(* IEC 61131-3 sources: KinematicsSimulation/crates/sim-opcua/examples/plc/twincat, 3 files *)

(* ---- sim_cycle.st ---- *)
(*
    A PLC cycle against the KinematicsSimulation link (sim-opcua), for TwinCAT 3 with TF6100 (library
    Tc3_PLCopen_OpcUa). Uses SIM_Access, SIM_MC_Power and SIM_MC_MoveAbsolute from sim_plcopen.st in this folder.

    NOT COMPILED: TwinCAT needs a Beckhoff account to download, so it was not built. The names were checked on
    14 November 2026 against Beckhoff Infosys (TF6100 TwinCAT 3 OPC UA Client, documentation 1.3.0 of 8 April 2026)
    and Beckhoff's TF6100_Samples on GitHub; what those do not settle is marked "CHECK".

    PRG_SimCycle:
      - connects with Basic256Sha256 SignAndEncrypt (or None, see bSecure), optionally with user name and password;
      - finds the namespace index from the URI 'urn:kinematics-simulation';
      - gets the node handles of the position and following error of one axis once and reads both every cycle,
        with the handles kept (one round trip per read; a read is started again as soon as the last one is done);
      - powers the axis (MC_Power), moves it with MC_MoveAbsolute, then writes a path and runs it
        (command.path, command.run_path) and waits until status.busy falls;
      - keeps the largest following error seen, switches off and disconnects.
    Run it in a task of 10 ms; sim-opcua then reports the task's write and read intervals (status.client_*).

    Data types as sim-opcua serves them (docs/plc.md, "Node ids and data types"): Double -> LREAL, Boolean -> BOOL,
    UInt16 -> UINT, Int32 -> DINT, UInt64 -> ULINT, String -> STRING. A PLC variable of another type (REAL for a
    Double) makes UA_Read fail with a type mismatch.
*)

FUNCTION_BLOCK SIM_CyclicRead
(* Reads one LREAL variable over and over through a node handle that is got once. *)
VAR_INPUT
    bEnable     : BOOL;
    hConnection : DWORD;
    nNamespace  : UINT;
    sNode       : STRING(255);
END_VAR
VAR_OUTPUT
    fValue  : LREAL;
    nReads  : UDINT;     (* reads done *)
    bError  : BOOL;
    nErrorID : DWORD;
END_VAR
VAR
    fbGetHandle : UA_NodeGetHandle;
    fbRead      : UA_Read;
    fbRelease   : UA_NodeReleaseHandle;
    stNodeID    : ST_UANodeID;
    stInfo      : ST_UANodeAdditionalInfo;
    hNode       : DWORD;
    nStep       : INT;
END_VAR

CASE nStep OF
0:  IF bEnable THEN
        stNodeID.nNamespaceIndex := nNamespace;
        stNodeID.sIdentifier := sNode;
        stNodeID.eIdentifierType := eUAIdentifierType_String;
        stInfo.eAttributeID := eUAAI_Value;   (* the Value attribute, 13 *)
        bError := FALSE; nErrorID := 0;
        nStep := 1;
    END_IF
1:  fbGetHandle(Execute := TRUE, ConnectionHdl := hConnection, NodeID := stNodeID);
    IF fbGetHandle.Done THEN
        hNode := fbGetHandle.NodeHdl; fbGetHandle(Execute := FALSE); nStep := 2;
    ELSIF fbGetHandle.Error THEN
        nErrorID := fbGetHandle.ErrorID; fbGetHandle(Execute := FALSE); bError := TRUE; nStep := 9;
    END_IF
2:  (* one read; once it is done the next starts in the same cycle, so a read that returns within a cycle runs
       every cycle *)
    fbRead(Execute := TRUE, ConnectionHdl := hConnection, NodeHdl := hNode, stNodeAddInfo := stInfo,
           cbData := SIZEOF(fValue), pVariable := ADR(fValue));
    IF fbRead.Done OR fbRead.Error THEN
        IF fbRead.Error THEN bError := TRUE; nErrorID := fbRead.ErrorID; ELSE nReads := nReads + 1; END_IF
        fbRead(Execute := FALSE);
        IF bEnable THEN
            fbRead(Execute := TRUE, ConnectionHdl := hConnection, NodeHdl := hNode, stNodeAddInfo := stInfo,
                   cbData := SIZEOF(fValue), pVariable := ADR(fValue));
        ELSE
            nStep := 3;
        END_IF
    END_IF
3:  fbRelease(Execute := TRUE, ConnectionHdl := hConnection, NodeHdl := hNode);
    IF fbRelease.Done OR fbRelease.Error THEN fbRelease(Execute := FALSE); nStep := 0; END_IF
9:  IF NOT bEnable THEN nStep := 0; END_IF
END_CASE
END_FUNCTION_BLOCK

PROGRAM PRG_SimCycle
VAR
    sServerUrl   : STRING(255) := 'opc.tcp://127.0.0.1:4840';   (* sim-opcua on the same PC *)
    bSecure      : BOOL := TRUE;                                 (* FALSE: SecurityPolicy None *)
    sUser        : STRING(63) := '';                             (* empty: anonymous; else as sim-opcua --user *)
    sPassword    : STRING(63) := '';
    sAxis        : STRING(31) := 'x';                            (* an axis id of the simulated machine *)
    fTarget      : LREAL := 0.4;                                 (* m, inside the axis range *)
    (* The path in the text of a path file, one piece per line ($N), one position per axis (here x and z of the
       T-gantry, which starts at x 0.1, z 0.35). *)
    sPath        : STRING(255) := 'line,0.4,0.25$Nline,0.1,0.25$Nline,0.1,0.35';
    (* sim-opcua counts every Read request: two reads a cycle show as intervals of half a cycle. FALSE reads the
       position alone, one request a cycle, so status.client_read_* give the task's cycle and jitter. *)
    bReadFollowingError : BOOL := TRUE;

    fbConnect    : UA_Connect;
    fbNamespace  : UA_GetNamespaceIndex;
    fbDisconnect : UA_Disconnect;
    stSession    : ST_UASessionConnectInfo;
    hConnection  : DWORD;
    nNamespace   : UINT;
    fbPower      : SIM_MC_Power;
    fbMove       : SIM_MC_MoveAbsolute;
    fbWrite      : SIM_Access;
    fbBusy       : SIM_Access;
    fbPosition   : SIM_CyclicRead;
    fbError      : SIM_CyclicRead;
    bTrue        : BOOL := TRUE;
    bBusy        : BOOL;
    bBusySeen    : BOOL;
    fLargestError : LREAL;   (* m, the largest following error read *)
    nStep        : INT;
END_VAR

CASE nStep OF
0:  stSession.sApplicationName := 'TwinCAT sim client';
    stSession.eTransportProfileUri := eUATransportProfileUri_UATcp;
    stSession.tSessionTimeout := T#60S;
    IF bSecure THEN
        (* TF6100 creates its own self-signed client certificate on its first start, in its PKI folder
           (%TcInstallDir%\3.1\Target\OpcUa\Client\PKI for client 2.x, %ProgramData%\Beckhoff\TF6100-OPC-UA\
           TcOpcUaClient\PKI for 1.x; Infosys "Application directories"). sim-opcua refuses it once and stores it in
           pki/rejected; move it to pki/trusted, or start sim-opcua with --trust-all while commissioning. TF6100
           likewise puts the server's certificate into its own rejected folder on the first attempt: move it to
           trusted there. *)
        stSession.eSecurityMode := eUASecurityMsgMode_Sign_Encrypt;
        stSession.eSecurityPolicyUri := eUASecurityPolicy_Basic256Sha256;
    ELSE
        stSession.eSecurityMode := eUASecurityMsgMode_None;
        stSession.eSecurityPolicyUri := eUASecurityPolicy_None;
    END_IF
    IF LEN(sUser) > 0 THEN
        stSession.stUserIdentTokenType.eUserIdentTokenType := eUAUITT_Username;
        stSession.stUserIdentTokenType.sTokenParam1 := sUser;
        stSession.stUserIdentTokenType.sTokenParam2 := sPassword;
    END_IF
    fbConnect(Execute := TRUE, ServerURL := sServerUrl, SessionConnectInfo := stSession, Timeout := T#5S);
    IF fbConnect.Done THEN hConnection := fbConnect.ConnectionHdl; fbConnect(Execute := FALSE); nStep := 10;
    ELSIF fbConnect.Error THEN fbConnect(Execute := FALSE); nStep := 900; END_IF
10: fbNamespace(Execute := TRUE, ConnectionHdl := hConnection, NamespaceUri := 'urn:kinematics-simulation', Timeout := T#5S);
    IF fbNamespace.Done THEN nNamespace := fbNamespace.NamespaceIndex; fbNamespace(Execute := FALSE); nStep := 20;
    ELSIF fbNamespace.Error THEN fbNamespace(Execute := FALSE); nStep := 900; END_IF
20: (* enable the drives *)
    fbPower.Enable := TRUE;
    IF fbPower.Status THEN nStep := 30; END_IF
30: (* MC_MoveAbsolute *)
    fbMove.Position := fTarget; fbMove.Velocity := 0.5; fbMove.Acceleration := 5.0; fbMove.Deceleration := 5.0;
    fbMove.Jerk := 100.0;
    fbMove.Execute := TRUE;
    IF fbMove.Done THEN fbMove.Execute := FALSE; nStep := 40;
    ELSIF fbMove.Error OR fbMove.CommandAborted THEN nStep := 900; END_IF
40: (* the path: its text, then command.run_path *)
    fbWrite(bExecute := FALSE);
    fbWrite(bExecute := TRUE, hConnection := hConnection, nNamespace := nNamespace, sNode := 'command.path',
            bWrite := TRUE, pData := ADR(sPath), cbData := LEN(sPath));
            (* CHECK: UA_Write documents cbData only as the size of the values to write; whether a STRING takes
               LEN (without the terminating null) or SIZEOF (the whole declared buffer) it does not say. *)
    nStep := 41;
41: fbWrite(bExecute := TRUE);
    IF fbWrite.bDone THEN nStep := 42; ELSIF fbWrite.bError THEN nStep := 900; END_IF
42: fbWrite(bExecute := FALSE);
    fbWrite(bExecute := TRUE, hConnection := hConnection, nNamespace := nNamespace, sNode := 'command.run_path',
            bWrite := TRUE, pData := ADR(bTrue), cbData := SIZEOF(bTrue));
    nStep := 43;
43: fbWrite(bExecute := TRUE);
    IF fbWrite.bDone THEN bBusySeen := FALSE; nStep := 50; ELSIF fbWrite.bError THEN nStep := 900; END_IF
50: (* poll status.busy until the path is over: it rises within a loop cycle or two and falls at the end *)
    fbBusy(bExecute := FALSE);
    fbBusy(bExecute := TRUE, hConnection := hConnection, nNamespace := nNamespace, sNode := 'status.busy',
           bWrite := FALSE, pData := ADR(bBusy), cbData := SIZEOF(bBusy));
    nStep := 51;
51: fbBusy(bExecute := TRUE);
    IF fbBusy.bDone THEN
        IF bBusy THEN bBusySeen := TRUE; nStep := 50;
        ELSIF bBusySeen THEN nStep := 60;
        ELSE nStep := 50; END_IF
    ELSIF fbBusy.bError THEN nStep := 900; END_IF
60: (* switch off and disconnect *)
    fbPower.Enable := FALSE;
    IF NOT fbPower.Status THEN nStep := 70; END_IF
70: fbDisconnect(Execute := TRUE, ConnectionHdl := hConnection, Timeout := T#5S);
    IF fbDisconnect.Done OR fbDisconnect.Error THEN fbDisconnect(Execute := FALSE); nStep := 100; END_IF
100: ; (* finished: fLargestError holds the largest following error *)
900: ; (* error: look at the blocks' ErrorID and at status.refused on the server *)
END_CASE

(* every cycle from the namespace on: position and following error of the axis *)
fbPosition(bEnable := nStep >= 20 AND nStep < 70, hConnection := hConnection, nNamespace := nNamespace,
           sNode := CONCAT(CONCAT('signal.axis.', sAxis), '.position'));
fbError(bEnable := bReadFollowingError AND nStep >= 20 AND nStep < 70, hConnection := hConnection, nNamespace := nNamespace,
        sNode := CONCAT(CONCAT('signal.axis.', sAxis), '.following_error'));
IF ABS(fbError.fValue) > fLargestError THEN fLargestError := ABS(fbError.fValue); END_IF

IF nStep >= 20 AND nStep < 70 THEN
    fbPower(hConnection := hConnection, nNamespace := nNamespace, sAxis := sAxis);
    fbMove(hConnection := hConnection, nNamespace := nNamespace, sAxis := sAxis);
END_IF
END_PROGRAM

(* ---- sim_plcopen.st ---- *)
(*
    PLCopen motion over OPC UA to the KinematicsSimulation link (sim-opcua), for TwinCAT 3.
    Library: Tc3_PLCopen_OpcUa (add it in the PLC project's References).

    NOT COMPILED: TwinCAT needs a Beckhoff account to download, so this file was not built. The names were checked
    on 14 November 2026 against Beckhoff Infosys (TF6100 TwinCAT 3 OPC UA Client, documentation 1.3.0 of
    8 April 2026) and Beckhoff's TF6100_Samples on GitHub.

    Structure:
      SIM_Access          one OPC UA read or write of one variable (get handle, read/write, release handle)
      SIM_Handshake       the PLCopen handshake of one function block on the simulator: inputs, Execute low,
                          wait for Done low, Execute high, poll Busy/Done/CommandAborted/Error/ErrorID
      SIM_MC_Power, SIM_MC_Home, SIM_MC_MoveAbsolute, SIM_MC_MoveRelative, SIM_MC_Stop, SIM_MC_Reset
                          thin wrappers with PLCopen inputs and outputs
      PRG_SimDemo         connect, power, home, move, stop, disconnect

    Node ids are strings in the namespace "urn:kinematics-simulation", e.g. 'axis.x.MoveAbsolute.Execute'.
    Getting a handle for every access keeps the code short and costs three round trips; cache the handles in
    production code.
*)

TYPE E_SimKind : (SIM_BOOL, SIM_LREAL, SIM_UINT); END_TYPE

FUNCTION_BLOCK SIM_Access
VAR_INPUT
    bExecute    : BOOL;            (* rising edge starts the access *)
    hConnection : DWORD;
    nNamespace  : UINT;
    sNode       : STRING(255);     (* e.g. 'axis.x.Power.Enable' *)
    bWrite      : BOOL;            (* TRUE: write the value at pData; FALSE: read into it *)
    pData       : PVOID;
    cbData      : UDINT;
END_VAR
VAR_OUTPUT
    bDone    : BOOL;
    bBusy    : BOOL;
    bError   : BOOL;
    nErrorID : DWORD;
END_VAR
VAR
    fbGetHandle : UA_NodeGetHandle;
    fbRead      : UA_Read;
    fbWrite     : UA_Write;
    fbRelease   : UA_NodeReleaseHandle;
    stNodeID    : ST_UANodeID;
    stInfo      : ST_UANodeAdditionalInfo;
    hNode       : DWORD;
    nStep       : INT;
    bLast       : BOOL;
END_VAR

IF bExecute AND NOT bLast THEN
    bDone := FALSE; bError := FALSE; nErrorID := 0; bBusy := TRUE;
    stNodeID.nNamespaceIndex := nNamespace;
    stNodeID.sIdentifier := sNode;
    stNodeID.eIdentifierType := eUAIdentifierType_String;
    stInfo.eAttributeID := eUAAI_Value;   (* the Value attribute, 13 *)
    nStep := 1;
END_IF
bLast := bExecute;

CASE nStep OF
1:  fbGetHandle(Execute := TRUE, ConnectionHdl := hConnection, NodeID := stNodeID);
    IF fbGetHandle.Done THEN
        hNode := fbGetHandle.NodeHdl;
        fbGetHandle(Execute := FALSE);
        nStep := 2;
    ELSIF fbGetHandle.Error THEN
        nErrorID := fbGetHandle.ErrorID;
        fbGetHandle(Execute := FALSE);
        bError := TRUE; bBusy := FALSE; nStep := 0;
    END_IF
2:  IF bWrite THEN
        fbWrite(Execute := TRUE, ConnectionHdl := hConnection, NodeHdl := hNode, stNodeAddInfo := stInfo,
                cbData := cbData, pVariable := pData);
        IF fbWrite.Done OR fbWrite.Error THEN
            bError := fbWrite.Error; nErrorID := fbWrite.ErrorID;
            fbWrite(Execute := FALSE);
            nStep := 3;
        END_IF
    ELSE
        fbRead(Execute := TRUE, ConnectionHdl := hConnection, NodeHdl := hNode, stNodeAddInfo := stInfo,
               cbData := cbData, pVariable := pData);
        IF fbRead.Done OR fbRead.Error THEN
            bError := fbRead.Error; nErrorID := fbRead.ErrorID;
            fbRead(Execute := FALSE);
            nStep := 3;
        END_IF
    END_IF
3:  fbRelease(Execute := TRUE, ConnectionHdl := hConnection, NodeHdl := hNode);
    IF fbRelease.Done OR fbRelease.Error THEN
        fbRelease(Execute := FALSE);
        bBusy := FALSE; bDone := NOT bError; nStep := 0;
    END_IF
END_CASE
END_FUNCTION_BLOCK

FUNCTION_BLOCK SIM_Handshake
VAR_INPUT
    Execute     : BOOL;
    hConnection : DWORD;
    nNamespace  : UINT;
    sAxis       : STRING(31);                  (* axis id, e.g. 'x' *)
    sFb         : STRING(31);                  (* 'Home', 'MoveAbsolute', 'MoveRelative', 'Stop', 'Reset' *)
    nParams     : INT;                         (* how many of the inputs below to write, 0..5 *)
    asParam     : ARRAY[1..5] OF STRING(31);   (* e.g. 'Position' *)
    afParam     : ARRAY[1..5] OF LREAL;
END_VAR
VAR_OUTPUT
    Done           : BOOL;
    Busy           : BOOL;
    Active         : BOOL;
    CommandAborted : BOOL;
    Error          : BOOL;
    ErrorID        : UINT;
END_VAR
VAR
    fbAccess  : SIM_Access;
    nPhase    : INT;      (* 0 idle, 1 inputs, 2 Execute low, 3 wait Done low, 4 Execute high, 5 poll, 6 finished *)
    nItem     : INT;
    bLast     : BOOL;
    bStarted  : BOOL;     (* fbAccess was triggered for the current item *)
    bValue    : BOOL;
    fValue    : LREAL;
    nValue    : UINT;
    bRemote   : ARRAY[1..4] OF BOOL;   (* Busy, Done, CommandAborted, Error as read *)
    sBase     : STRING(80);
END_VAR

IF Execute AND NOT bLast THEN
    Done := FALSE; Busy := TRUE; Active := FALSE; CommandAborted := FALSE; Error := FALSE; ErrorID := 0;
    sBase := CONCAT(CONCAT(CONCAT('axis.', sAxis), '.'), CONCAT(sFb, '.'));
    IF nParams > 0 THEN nPhase := 1; ELSE nPhase := 2; END_IF
    nItem := 1; bStarted := FALSE;
ELSIF NOT Execute AND bLast THEN
    (* PLCopen: the outputs fall with Execute; the simulator's Execute goes low with it *)
    Done := FALSE; CommandAborted := FALSE; Error := FALSE; ErrorID := 0;
    IF NOT Busy THEN nPhase := 2; nItem := 1; bStarted := FALSE; END_IF
END_IF
bLast := Execute;

IF nPhase > 0 AND nPhase < 6 THEN
    IF NOT bStarted THEN
        (* the access of this phase and item *)
        fbAccess.hConnection := hConnection;
        fbAccess.nNamespace := nNamespace;
        CASE nPhase OF
        1:  fbAccess.sNode := CONCAT(sBase, asParam[nItem]); fValue := afParam[nItem];
            fbAccess.bWrite := TRUE; fbAccess.pData := ADR(fValue); fbAccess.cbData := SIZEOF(fValue);
        2, 4:
            fbAccess.sNode := CONCAT(sBase, 'Execute'); bValue := nPhase = 4;
            fbAccess.bWrite := TRUE; fbAccess.pData := ADR(bValue); fbAccess.cbData := SIZEOF(bValue);
        3:  fbAccess.sNode := CONCAT(sBase, 'Done');
            fbAccess.bWrite := FALSE; fbAccess.pData := ADR(bValue); fbAccess.cbData := SIZEOF(bValue);
        5:  IF nItem <= 4 THEN
                CASE nItem OF
                1: fbAccess.sNode := CONCAT(sBase, 'Busy');
                2: fbAccess.sNode := CONCAT(sBase, 'Done');
                3: fbAccess.sNode := CONCAT(sBase, 'CommandAborted');
                4: fbAccess.sNode := CONCAT(sBase, 'Error');
                END_CASE
                fbAccess.pData := ADR(bValue); fbAccess.cbData := SIZEOF(bValue);
            ELSE
                fbAccess.sNode := CONCAT(sBase, 'ErrorID');
                fbAccess.pData := ADR(nValue); fbAccess.cbData := SIZEOF(nValue);
            END_IF
            fbAccess.bWrite := FALSE;
        END_CASE
        fbAccess(bExecute := FALSE);
        fbAccess(bExecute := TRUE);
        bStarted := TRUE;
    ELSE
        fbAccess(bExecute := TRUE);
    END_IF

    IF fbAccess.bError THEN
        Error := TRUE; ErrorID := 16#FFFF; Busy := FALSE; nPhase := 6;   (* the OPC UA access failed *)
    ELSIF fbAccess.bDone THEN
        bStarted := FALSE;
        CASE nPhase OF
        1:  nItem := nItem + 1;
            IF nItem > nParams THEN nPhase := 2; nItem := 1; END_IF
        2:  IF Busy THEN nPhase := 3; ELSE nPhase := 0; END_IF   (* after the falling edge: done *)
        3:  IF NOT bValue THEN nPhase := 4; END_IF                (* outputs are published once a cycle *)
        4:  nPhase := 5; nItem := 1;
        5:  IF nItem <= 4 THEN
                bRemote[nItem] := bValue;
                nItem := nItem + 1;
            ELSE
                ErrorID := nValue;
                Active := bRemote[1];
                IF bRemote[2] OR bRemote[3] OR bRemote[4] THEN
                    Done := bRemote[2] AND Execute;
                    CommandAborted := bRemote[3] AND Execute;
                    Error := bRemote[4] AND Execute;
                    Busy := FALSE; Active := FALSE;
                    nPhase := 6;
                END_IF
                nItem := 1;
            END_IF
        END_CASE
    END_IF
END_IF
END_FUNCTION_BLOCK

FUNCTION_BLOCK SIM_MC_Power
VAR_INPUT
    Enable      : BOOL;
    hConnection : DWORD;
    nNamespace  : UINT;
    sAxis       : STRING(31);
END_VAR
VAR_OUTPUT
    Status : BOOL;
    Valid  : BOOL;
    Error  : BOOL;
END_VAR
VAR
    fbAccess : SIM_Access;
    nStep    : INT;
    bWritten : BOOL;   (* the Enable last written *)
    bValue   : BOOL;
    bFirst   : BOOL := TRUE;
END_VAR

(* writes Enable when it changes, otherwise reads Power.Status *)
CASE nStep OF
0:  fbAccess.hConnection := hConnection; fbAccess.nNamespace := nNamespace;
    IF bFirst OR Enable <> bWritten THEN
        bValue := Enable; bWritten := Enable; bFirst := FALSE;
        fbAccess.sNode := CONCAT(CONCAT('axis.', sAxis), '.Power.Enable');
        fbAccess.bWrite := TRUE;
    ELSE
        fbAccess.sNode := CONCAT(CONCAT('axis.', sAxis), '.Power.Status');
        fbAccess.bWrite := FALSE;
    END_IF
    fbAccess.pData := ADR(bValue); fbAccess.cbData := SIZEOF(bValue);
    fbAccess(bExecute := FALSE);
    fbAccess(bExecute := TRUE);
    nStep := 1;
1:  fbAccess(bExecute := TRUE);
    IF fbAccess.bDone OR fbAccess.bError THEN
        Error := fbAccess.bError;
        IF fbAccess.bDone AND NOT fbAccess.bWrite THEN Status := bValue; END_IF
        Valid := Status AND NOT Error;
        nStep := 0;
    END_IF
END_CASE
END_FUNCTION_BLOCK

FUNCTION_BLOCK SIM_MC_Home
VAR_INPUT
    Execute : BOOL; hConnection : DWORD; nNamespace : UINT; sAxis : STRING(31);
END_VAR
VAR_OUTPUT
    Done : BOOL; Busy : BOOL; Active : BOOL; CommandAborted : BOOL; Error : BOOL; ErrorID : UINT;
END_VAR
VAR
    fbCall : SIM_Handshake;
END_VAR
fbCall(Execute := Execute, hConnection := hConnection, nNamespace := nNamespace, sAxis := sAxis, sFb := 'Home', nParams := 0);
Done := fbCall.Done; Busy := fbCall.Busy; Active := fbCall.Active;
CommandAborted := fbCall.CommandAborted; Error := fbCall.Error; ErrorID := fbCall.ErrorID;
END_FUNCTION_BLOCK

FUNCTION_BLOCK SIM_MC_MoveAbsolute
VAR_INPUT
    Execute : BOOL; hConnection : DWORD; nNamespace : UINT; sAxis : STRING(31);
    Position : LREAL; Velocity : LREAL; Acceleration : LREAL; Deceleration : LREAL; Jerk : LREAL;
END_VAR
VAR_OUTPUT
    Done : BOOL; Busy : BOOL; Active : BOOL; CommandAborted : BOOL; Error : BOOL; ErrorID : UINT;
END_VAR
VAR
    fbCall : SIM_Handshake;
END_VAR
fbCall.asParam[1] := 'Position';     fbCall.afParam[1] := Position;
fbCall.asParam[2] := 'Velocity';     fbCall.afParam[2] := Velocity;
fbCall.asParam[3] := 'Acceleration'; fbCall.afParam[3] := Acceleration;
fbCall.asParam[4] := 'Deceleration'; fbCall.afParam[4] := Deceleration;
fbCall.asParam[5] := 'Jerk';         fbCall.afParam[5] := Jerk;
fbCall(Execute := Execute, hConnection := hConnection, nNamespace := nNamespace, sAxis := sAxis, sFb := 'MoveAbsolute', nParams := 5);
Done := fbCall.Done; Busy := fbCall.Busy; Active := fbCall.Active;
CommandAborted := fbCall.CommandAborted; Error := fbCall.Error; ErrorID := fbCall.ErrorID;
END_FUNCTION_BLOCK

FUNCTION_BLOCK SIM_MC_MoveRelative
VAR_INPUT
    Execute : BOOL; hConnection : DWORD; nNamespace : UINT; sAxis : STRING(31);
    Distance : LREAL; Velocity : LREAL; Acceleration : LREAL; Deceleration : LREAL; Jerk : LREAL;
END_VAR
VAR_OUTPUT
    Done : BOOL; Busy : BOOL; Active : BOOL; CommandAborted : BOOL; Error : BOOL; ErrorID : UINT;
END_VAR
VAR
    fbCall : SIM_Handshake;
END_VAR
fbCall.asParam[1] := 'Distance';     fbCall.afParam[1] := Distance;
fbCall.asParam[2] := 'Velocity';     fbCall.afParam[2] := Velocity;
fbCall.asParam[3] := 'Acceleration'; fbCall.afParam[3] := Acceleration;
fbCall.asParam[4] := 'Deceleration'; fbCall.afParam[4] := Deceleration;
fbCall.asParam[5] := 'Jerk';         fbCall.afParam[5] := Jerk;
fbCall(Execute := Execute, hConnection := hConnection, nNamespace := nNamespace, sAxis := sAxis, sFb := 'MoveRelative', nParams := 5);
Done := fbCall.Done; Busy := fbCall.Busy; Active := fbCall.Active;
CommandAborted := fbCall.CommandAborted; Error := fbCall.Error; ErrorID := fbCall.ErrorID;
END_FUNCTION_BLOCK

FUNCTION_BLOCK SIM_MC_Stop
VAR_INPUT
    Execute : BOOL; hConnection : DWORD; nNamespace : UINT; sAxis : STRING(31);
    Deceleration : LREAL;
END_VAR
VAR_OUTPUT
    Done : BOOL; Busy : BOOL; Active : BOOL; CommandAborted : BOOL; Error : BOOL; ErrorID : UINT;
END_VAR
VAR
    fbCall : SIM_Handshake;
END_VAR
fbCall.asParam[1] := 'Deceleration'; fbCall.afParam[1] := Deceleration;
fbCall(Execute := Execute, hConnection := hConnection, nNamespace := nNamespace, sAxis := sAxis, sFb := 'Stop', nParams := 1);
Done := fbCall.Done; Busy := fbCall.Busy; Active := fbCall.Active;
CommandAborted := fbCall.CommandAborted; Error := fbCall.Error; ErrorID := fbCall.ErrorID;
END_FUNCTION_BLOCK

FUNCTION_BLOCK SIM_MC_Reset
VAR_INPUT
    Execute : BOOL; hConnection : DWORD; nNamespace : UINT; sAxis : STRING(31);
END_VAR
VAR_OUTPUT
    Done : BOOL; Busy : BOOL; Error : BOOL; ErrorID : UINT;
END_VAR
VAR
    fbCall : SIM_Handshake;
END_VAR
fbCall(Execute := Execute, hConnection := hConnection, nNamespace := nNamespace, sAxis := sAxis, sFb := 'Reset', nParams := 0);
Done := fbCall.Done; Busy := fbCall.Busy; Error := fbCall.Error; ErrorID := fbCall.ErrorID;
END_FUNCTION_BLOCK

PROGRAM PRG_SimDemo
VAR
    fbConnect    : UA_Connect;
    fbNamespace  : UA_GetNamespaceIndex;
    fbDisconnect : UA_Disconnect;
    stSession    : ST_UASessionConnectInfo;
    hConnection  : DWORD;
    nNamespace   : UINT;
    fbPower      : SIM_MC_Power;
    fbHome       : SIM_MC_Home;
    fbMove       : SIM_MC_MoveAbsolute;
    fbStop       : SIM_MC_Stop;
    tonMoving    : TON;
    nStep        : INT;
    sAxis        : STRING(31) := 'x';    (* an axis id of the simulated machine *)
END_VAR

CASE nStep OF
0:  (* connect without security; the link offers SecurityPolicy None with anonymous login *)
    stSession.sApplicationName := 'TwinCAT sim client';
    stSession.eSecurityMode := eUASecurityMsgMode_None;
    stSession.eSecurityPolicyUri := eUASecurityPolicy_None;
    stSession.eTransportProfileUri := eUATransportProfileUri_UATcp;
    stSession.tSessionTimeout := T#60S;
    fbConnect(Execute := TRUE, ServerURL := 'opc.tcp://192.168.0.10:4840', SessionConnectInfo := stSession, Timeout := T#5S);
    IF fbConnect.Done THEN hConnection := fbConnect.ConnectionHdl; fbConnect(Execute := FALSE); nStep := 10;
    ELSIF fbConnect.Error THEN fbConnect(Execute := FALSE); nStep := 900; END_IF
10: fbNamespace(Execute := TRUE, ConnectionHdl := hConnection, NamespaceUri := 'urn:kinematics-simulation', Timeout := T#5S);
    IF fbNamespace.Done THEN nNamespace := fbNamespace.NamespaceIndex; fbNamespace(Execute := FALSE); nStep := 20;
    ELSIF fbNamespace.Error THEN fbNamespace(Execute := FALSE); nStep := 900; END_IF
20: (* power on *)
    fbPower.Enable := TRUE;
    IF fbPower.Status THEN nStep := 30; END_IF
30: (* home *)
    fbHome.Execute := TRUE;
    IF fbHome.Done THEN fbHome.Execute := FALSE; nStep := 40;
    ELSIF fbHome.Error THEN nStep := 900; END_IF
40: (* move absolute, stopped after 0.5 s *)
    fbMove.Position := 0.6; fbMove.Velocity := 0.5; fbMove.Acceleration := 5.0; fbMove.Deceleration := 5.0; fbMove.Jerk := 100.0;
    fbMove.Execute := TRUE;
    tonMoving(IN := fbMove.Busy, PT := T#500MS);
    IF tonMoving.Q OR fbMove.Done THEN nStep := 50;
    ELSIF fbMove.Error THEN nStep := 900; END_IF
50: fbStop.Deceleration := 2.0;
    fbStop.Execute := TRUE;
    IF fbStop.Done THEN fbStop.Execute := FALSE; fbMove.Execute := FALSE; nStep := 60;
    ELSIF fbStop.Error THEN nStep := 900; END_IF
60: (* power off and disconnect *)
    fbPower.Enable := FALSE;
    IF NOT fbPower.Status THEN nStep := 70; END_IF
70: fbDisconnect(Execute := TRUE, ConnectionHdl := hConnection, Timeout := T#5S);
    IF fbDisconnect.Done OR fbDisconnect.Error THEN fbDisconnect(Execute := FALSE); nStep := 100; END_IF
100: ; (* finished *)
900: ; (* error: look at the blocks' ErrorID *)
END_CASE

IF nStep >= 20 AND nStep < 70 THEN
    fbPower(hConnection := hConnection, nNamespace := nNamespace, sAxis := sAxis);
    fbHome(hConnection := hConnection, nNamespace := nNamespace, sAxis := sAxis);
    fbMove(hConnection := hConnection, nNamespace := nNamespace, sAxis := sAxis);
    fbStop(hConnection := hConnection, nNamespace := nNamespace, sAxis := sAxis);
END_IF
END_PROGRAM

(* ---- sim_sync.st ---- *)
(*
    PLCopen synchronised motion over OPC UA to the KinematicsSimulation link (sim-opcua), for TwinCAT 3:
    MC_GearIn, MC_GearOut, MC_CamIn and MC_CamOut on a slave axis, its master another axis of the machine.
    Library: Tc3_PLCopen_OpcUa. Needs SIM_Access and SIM_Handshake from sim_plcopen.st in the same project.

    NOT COMPILED: TwinCAT needs a Beckhoff account to download, so this file was not built. It uses only the blocks
    of sim_plcopen.st (whose names were checked there) and plain IEC 61131-3. CHECK: the size TF6100's UA_Write
    takes for a STRING (here LEN + 1, the text and its terminating zero); the link reads the text up to its end.

    Structure:
      SIM_WriteText        one write of a text input (GearIn.Master, CamIn.Master, CamIn.Table)
      SIM_SyncHandshake    the handshake of MC_GearIn or MC_CamIn: inputs and texts, Execute low, Execute high, then
                           poll Busy, InGear/InSync, CommandAborted, Error and ErrorID for as long as the block is busy:
                           unlike a move it stays busy while the slave is coupled
      SIM_MC_GearIn, SIM_MC_CamIn, SIM_MC_GearOut, SIM_MC_CamOut   thin wrappers with PLCopen inputs and outputs
      PRG_SimSyncDemo      x moves, y gears in at 2:1, gears out, cams in on a 3-4-5 table, cams out, stops

    The master is named by its axis id ('x'); an empty CamIn.Master with CamTableID 1 runs the slave on the machine's
    own electronic cam and its virtual master (the crank and cam machines). See docs/plc.md.
*)

FUNCTION_BLOCK SIM_WriteText
VAR_INPUT
    bExecute    : BOOL;
    hConnection : DWORD;
    nNamespace  : UINT;
    sNode       : STRING(255);
    sText       : STRING(1023);
END_VAR
VAR_OUTPUT
    bDone : BOOL; bBusy : BOOL; bError : BOOL; nErrorID : DWORD;
END_VAR
VAR
    fbAccess : SIM_Access;
END_VAR
fbAccess(bExecute := bExecute, hConnection := hConnection, nNamespace := nNamespace, sNode := sNode, bWrite := TRUE,
         pData := ADR(sText), cbData := INT_TO_UDINT(LEN(sText)) + 1);
bDone := fbAccess.bDone; bBusy := fbAccess.bBusy; bError := fbAccess.bError; nErrorID := fbAccess.nErrorID;
END_FUNCTION_BLOCK

FUNCTION_BLOCK SIM_SyncHandshake
VAR_INPUT
    Execute     : BOOL;
    hConnection : DWORD;
    nNamespace  : UINT;
    sAxis       : STRING(31);                  (* the slave's axis id *)
    sFb         : STRING(31);                  (* 'GearIn' or 'CamIn' *)
    sMaster     : STRING(31);                  (* the master's axis id; '' for the machine's virtual cam master *)
    sTable      : STRING(1023);                (* CamIn only: the cam table, '' to leave it as it is *)
    nParams     : INT;                         (* 0..6 *)
    asParam     : ARRAY[1..6] OF STRING(31);
    afParam     : ARRAY[1..6] OF LREAL;
END_VAR
VAR_OUTPUT
    InSync         : BOOL;     (* InGear of MC_GearIn, InSync of MC_CamIn *)
    Busy           : BOOL;
    Active         : BOOL;
    CommandAborted : BOOL;
    Error          : BOOL;
    ErrorID        : UINT;
END_VAR
VAR
    fbAccess : SIM_Access;
    fbText   : SIM_WriteText;
    nPhase   : INT;      (* 0 idle, 1 inputs, 2 Master, 3 Table, 4 Execute low, 5 Execute high, 6 poll, 7 finished *)
    nItem    : INT;
    bLast    : BOOL;
    bStarted : BOOL;
    bValue   : BOOL;
    fValue   : LREAL;
    nValue   : UINT;
    bRemote  : ARRAY[1..4] OF BOOL;   (* Busy, InGear/InSync, CommandAborted, Error as read *)
    sBase    : STRING(80);
    sSync    : STRING(31);
END_VAR

IF Execute AND NOT bLast THEN
    InSync := FALSE; Busy := TRUE; Active := FALSE; CommandAborted := FALSE; Error := FALSE; ErrorID := 0;
    sBase := CONCAT(CONCAT(CONCAT('axis.', sAxis), '.'), CONCAT(sFb, '.'));
    IF sFb = 'GearIn' THEN sSync := 'InGear'; ELSE sSync := 'InSync'; END_IF
    IF nParams > 0 THEN nPhase := 1; ELSE nPhase := 2; END_IF
    nItem := 1; bStarted := FALSE;
ELSIF NOT Execute AND bLast THEN
    (* the outputs fall with Execute; a coupled block stays coupled until GearOut/CamOut or another block *)
    InSync := FALSE; CommandAborted := FALSE; Error := FALSE; ErrorID := 0;
    nPhase := 4; bStarted := FALSE;
END_IF
bLast := Execute;

IF nPhase = 2 OR nPhase = 3 THEN
    (* the texts: the master, then (CamIn) the table *)
    IF nPhase = 3 AND (sFb <> 'CamIn' OR LEN(sTable) = 0) THEN
        nPhase := 4;
    ELSE
        IF NOT bStarted THEN
            fbText.hConnection := hConnection; fbText.nNamespace := nNamespace;
            IF nPhase = 2 THEN
                fbText.sNode := CONCAT(sBase, 'Master'); fbText.sText := sMaster;
            ELSE
                fbText.sNode := CONCAT(sBase, 'Table'); fbText.sText := sTable;
            END_IF
            fbText(bExecute := FALSE);
            bStarted := TRUE;
        END_IF
        fbText(bExecute := TRUE);
        IF fbText.bError THEN
            Error := TRUE; ErrorID := 16#FFFF; Busy := FALSE; nPhase := 7;
        ELSIF fbText.bDone THEN
            bStarted := FALSE; nPhase := nPhase + 1;
        END_IF
    END_IF
ELSIF nPhase > 0 AND nPhase < 7 THEN
    IF NOT bStarted THEN
        fbAccess.hConnection := hConnection;
        fbAccess.nNamespace := nNamespace;
        CASE nPhase OF
        1:  fbAccess.sNode := CONCAT(sBase, asParam[nItem]); fValue := afParam[nItem];
            fbAccess.bWrite := TRUE; fbAccess.pData := ADR(fValue); fbAccess.cbData := SIZEOF(fValue);
        4, 5:
            fbAccess.sNode := CONCAT(sBase, 'Execute'); bValue := nPhase = 5 AND Execute;
            fbAccess.bWrite := TRUE; fbAccess.pData := ADR(bValue); fbAccess.cbData := SIZEOF(bValue);
        6:  IF nItem <= 4 THEN
                CASE nItem OF
                1: fbAccess.sNode := CONCAT(sBase, 'Busy');
                2: fbAccess.sNode := CONCAT(sBase, sSync);
                3: fbAccess.sNode := CONCAT(sBase, 'CommandAborted');
                4: fbAccess.sNode := CONCAT(sBase, 'Error');
                END_CASE
                fbAccess.pData := ADR(bValue); fbAccess.cbData := SIZEOF(bValue);
            ELSE
                fbAccess.sNode := CONCAT(sBase, 'ErrorID');
                fbAccess.pData := ADR(nValue); fbAccess.cbData := SIZEOF(nValue);
            END_IF
            fbAccess.bWrite := FALSE;
        END_CASE
        fbAccess(bExecute := FALSE);
        fbAccess(bExecute := TRUE);
        bStarted := TRUE;
    ELSE
        fbAccess(bExecute := TRUE);
    END_IF

    IF fbAccess.bError THEN
        Error := TRUE; ErrorID := 16#FFFF; Busy := FALSE; nPhase := 7;   (* the OPC UA access failed *)
    ELSIF fbAccess.bDone THEN
        bStarted := FALSE;
        CASE nPhase OF
        1:  nItem := nItem + 1;
            IF nItem > nParams THEN nPhase := 2; nItem := 1; END_IF
        4:  IF Execute THEN nPhase := 5; ELSE nPhase := 0; Busy := FALSE; Active := FALSE; END_IF
        5:  nPhase := 6; nItem := 1;
        6:  IF nItem <= 4 THEN
                bRemote[nItem] := bValue;
                nItem := nItem + 1;
            ELSE
                ErrorID := nValue;
                Busy := bRemote[1]; Active := bRemote[1];
                InSync := bRemote[2] AND Execute;
                CommandAborted := bRemote[3] AND Execute;
                Error := bRemote[4] AND Execute;
                (* coupled, the block stays busy: poll on; it is over once it is no longer busy *)
                IF NOT Busy THEN nPhase := 7; END_IF
                nItem := 1;
            END_IF
        END_CASE
    END_IF
END_IF
END_FUNCTION_BLOCK

FUNCTION_BLOCK SIM_MC_GearIn
VAR_INPUT
    Execute : BOOL; hConnection : DWORD; nNamespace : UINT;
    sMaster : STRING(31); sSlave : STRING(31);
    RatioNumerator : LREAL; RatioDenominator : LREAL; Acceleration : LREAL; Deceleration : LREAL; Jerk : LREAL;
END_VAR
VAR_OUTPUT
    InGear : BOOL; Busy : BOOL; Active : BOOL; CommandAborted : BOOL; Error : BOOL; ErrorID : UINT;
END_VAR
VAR
    fbCall : SIM_SyncHandshake;
END_VAR
fbCall.asParam[1] := 'RatioNumerator';   fbCall.afParam[1] := RatioNumerator;
fbCall.asParam[2] := 'RatioDenominator'; fbCall.afParam[2] := RatioDenominator;
fbCall.asParam[3] := 'Acceleration';     fbCall.afParam[3] := Acceleration;
fbCall.asParam[4] := 'Deceleration';     fbCall.afParam[4] := Deceleration;
fbCall.asParam[5] := 'Jerk';             fbCall.afParam[5] := Jerk;
fbCall(Execute := Execute, hConnection := hConnection, nNamespace := nNamespace, sAxis := sSlave, sFb := 'GearIn',
       sMaster := sMaster, sTable := '', nParams := 5);
InGear := fbCall.InSync; Busy := fbCall.Busy; Active := fbCall.Active;
CommandAborted := fbCall.CommandAborted; Error := fbCall.Error; ErrorID := fbCall.ErrorID;
END_FUNCTION_BLOCK

FUNCTION_BLOCK SIM_MC_CamIn
VAR_INPUT
    Execute : BOOL; hConnection : DWORD; nNamespace : UINT;
    sMaster : STRING(31); sSlave : STRING(31);
    MasterOffset : LREAL; SlaveOffset : LREAL; MasterScaling : LREAL := 1.0; SlaveScaling : LREAL := 1.0;
    StartMode : LREAL := 1.0;    (* 0 absolute, 1 relative *)
    CamTableID : LREAL;          (* 0 the table below, 1 the machine's own cam *)
    sTable : STRING(1023);       (* lines 'master span, slave rise, law' or 'master, slave[, slope]' *)
END_VAR
VAR_OUTPUT
    InSync : BOOL; Busy : BOOL; Active : BOOL; CommandAborted : BOOL; Error : BOOL; ErrorID : UINT;
END_VAR
VAR
    fbCall : SIM_SyncHandshake;
END_VAR
fbCall.asParam[1] := 'MasterOffset';  fbCall.afParam[1] := MasterOffset;
fbCall.asParam[2] := 'SlaveOffset';   fbCall.afParam[2] := SlaveOffset;
fbCall.asParam[3] := 'MasterScaling'; fbCall.afParam[3] := MasterScaling;
fbCall.asParam[4] := 'SlaveScaling';  fbCall.afParam[4] := SlaveScaling;
fbCall.asParam[5] := 'StartMode';     fbCall.afParam[5] := StartMode;
fbCall.asParam[6] := 'CamTableID';    fbCall.afParam[6] := CamTableID;
fbCall(Execute := Execute, hConnection := hConnection, nNamespace := nNamespace, sAxis := sSlave, sFb := 'CamIn',
       sMaster := sMaster, sTable := sTable, nParams := 6);
InSync := fbCall.InSync; Busy := fbCall.Busy; Active := fbCall.Active;
CommandAborted := fbCall.CommandAborted; Error := fbCall.Error; ErrorID := fbCall.ErrorID;
END_FUNCTION_BLOCK

FUNCTION_BLOCK SIM_MC_GearOut
VAR_INPUT
    Execute : BOOL; hConnection : DWORD; nNamespace : UINT; sSlave : STRING(31);
END_VAR
VAR_OUTPUT
    Done : BOOL; Busy : BOOL; Error : BOOL; ErrorID : UINT;
END_VAR
VAR
    fbCall : SIM_Handshake;
END_VAR
fbCall(Execute := Execute, hConnection := hConnection, nNamespace := nNamespace, sAxis := sSlave, sFb := 'GearOut', nParams := 0);
Done := fbCall.Done; Busy := fbCall.Busy; Error := fbCall.Error; ErrorID := fbCall.ErrorID;
END_FUNCTION_BLOCK

FUNCTION_BLOCK SIM_MC_CamOut
VAR_INPUT
    Execute : BOOL; hConnection : DWORD; nNamespace : UINT; sSlave : STRING(31);
END_VAR
VAR_OUTPUT
    Done : BOOL; Busy : BOOL; Error : BOOL; ErrorID : UINT;
END_VAR
VAR
    fbCall : SIM_Handshake;
END_VAR
fbCall(Execute := Execute, hConnection := hConnection, nNamespace := nNamespace, sAxis := sSlave, sFb := 'CamOut', nParams := 0);
Done := fbCall.Done; Busy := fbCall.Busy; Error := fbCall.Error; ErrorID := fbCall.ErrorID;
END_FUNCTION_BLOCK

PROGRAM PRG_SimSyncDemo
VAR
    fbConnect    : UA_Connect;
    fbNamespace  : UA_GetNamespaceIndex;
    fbDisconnect : UA_Disconnect;
    stSession    : ST_UASessionConnectInfo;
    hConnection  : DWORD;
    nNamespace   : UINT;
    fbPowerX     : SIM_MC_Power;
    fbPowerY     : SIM_MC_Power;
    fbMoveX      : SIM_MC_MoveAbsolute;
    fbGearIn     : SIM_MC_GearIn;
    fbGearOut    : SIM_MC_GearOut;
    fbCamIn      : SIM_MC_CamIn;
    fbCamOut     : SIM_MC_CamOut;
    fbStopY      : SIM_MC_Stop;
    tonGeared    : TON;
    nStep        : INT;
    sMaster      : STRING(31) := 'x';    (* axis ids of the simulated machine: a two-axis gantry *)
    sSlave       : STRING(31) := 'y';
END_VAR

CASE nStep OF
0:  stSession.sApplicationName := 'TwinCAT sim client';
    stSession.eSecurityMode := eUASecurityMsgMode_None;
    stSession.eSecurityPolicyUri := eUASecurityPolicy_None;
    stSession.eTransportProfileUri := eUATransportProfileUri_UATcp;
    stSession.tSessionTimeout := T#60S;
    fbConnect(Execute := TRUE, ServerURL := 'opc.tcp://192.168.0.10:4840', SessionConnectInfo := stSession, Timeout := T#5S);
    IF fbConnect.Done THEN hConnection := fbConnect.ConnectionHdl; fbConnect(Execute := FALSE); nStep := 10;
    ELSIF fbConnect.Error THEN fbConnect(Execute := FALSE); nStep := 900; END_IF
10: fbNamespace(Execute := TRUE, ConnectionHdl := hConnection, NamespaceUri := 'urn:kinematics-simulation', Timeout := T#5S);
    IF fbNamespace.Done THEN nNamespace := fbNamespace.NamespaceIndex; fbNamespace(Execute := FALSE); nStep := 20;
    ELSIF fbNamespace.Error THEN fbNamespace(Execute := FALSE); nStep := 900; END_IF
20: fbPowerX.Enable := TRUE; fbPowerY.Enable := TRUE;
    IF fbPowerX.Status AND fbPowerY.Status THEN nStep := 30; END_IF
30: (* the master runs slowly over its stroke *)
    fbMoveX.Position := 0.9; fbMoveX.Velocity := 0.05; fbMoveX.Acceleration := 1.0; fbMoveX.Deceleration := 1.0;
    fbMoveX.Jerk := 100.0; fbMoveX.Execute := TRUE;
    IF fbMoveX.Busy THEN nStep := 40; ELSIF fbMoveX.Error THEN nStep := 900; END_IF
40: (* y gears in at 2:1 *)
    fbGearIn.RatioNumerator := 2.0; fbGearIn.RatioDenominator := 1.0;
    fbGearIn.Acceleration := 1.0; fbGearIn.Deceleration := 1.0; fbGearIn.Jerk := 100.0;
    fbGearIn.Execute := TRUE;
    tonGeared(IN := fbGearIn.InGear, PT := T#1S);
    IF tonGeared.Q THEN nStep := 50; ELSIF fbGearIn.Error OR fbGearIn.CommandAborted THEN nStep := 900; END_IF
50: fbGearOut.Execute := TRUE;
    IF fbGearOut.Done THEN fbGearOut.Execute := FALSE; fbGearIn.Execute := FALSE; nStep := 60;
    ELSIF fbGearOut.Error THEN nStep := 900; END_IF
60: (* y cams in, relative, on a 3-4-5 rise of 20 mm over 0.1 m of x and back *)
    fbCamIn.sTable := '0.1, 0.02, 3-4-5$N0.1, -0.02, 3-4-5';
    fbCamIn.StartMode := 1.0; fbCamIn.CamTableID := 0.0;
    fbCamIn.Execute := TRUE;
    IF fbCamIn.InSync THEN nStep := 70; ELSIF fbCamIn.Error THEN nStep := 900; END_IF
70: IF NOT fbMoveX.Busy THEN nStep := 80; END_IF   (* x has arrived; y stands on its cam *)
80: fbCamOut.Execute := TRUE;
    IF fbCamOut.Done THEN fbCamOut.Execute := FALSE; fbCamIn.Execute := FALSE; nStep := 90;
    ELSIF fbCamOut.Error THEN nStep := 900; END_IF
90: fbStopY.Deceleration := 1.0; fbStopY.Execute := TRUE;
    IF fbStopY.Done THEN fbStopY.Execute := FALSE; fbMoveX.Execute := FALSE; nStep := 95;
    ELSIF fbStopY.Error THEN nStep := 900; END_IF
95: fbPowerX.Enable := FALSE; fbPowerY.Enable := FALSE;
    IF NOT fbPowerX.Status AND NOT fbPowerY.Status THEN nStep := 99; END_IF
99: fbDisconnect(Execute := TRUE, ConnectionHdl := hConnection, Timeout := T#5S);
    IF fbDisconnect.Done OR fbDisconnect.Error THEN fbDisconnect(Execute := FALSE); nStep := 100; END_IF
100: ; (* finished *)
900: ; (* error: look at the blocks' ErrorID *)
END_CASE

IF nStep >= 20 AND nStep < 99 THEN
    fbPowerX(hConnection := hConnection, nNamespace := nNamespace, sAxis := sMaster);
    fbPowerY(hConnection := hConnection, nNamespace := nNamespace, sAxis := sSlave);
    fbMoveX(hConnection := hConnection, nNamespace := nNamespace, sAxis := sMaster);
    fbGearIn(hConnection := hConnection, nNamespace := nNamespace, sMaster := sMaster, sSlave := sSlave);
    fbGearOut(hConnection := hConnection, nNamespace := nNamespace, sSlave := sSlave);
    fbCamIn(hConnection := hConnection, nNamespace := nNamespace, sMaster := sMaster, sSlave := sSlave);
    fbCamOut(hConnection := hConnection, nNamespace := nNamespace, sSlave := sSlave);
    fbStopY(hConnection := hConnection, nNamespace := nNamespace, sAxis := sSlave);
END_IF
END_PROGRAM
